(*
SPDX-FileCopyrightText: © 2026 Oleksandr Tiutyk <trofimich@gmail.com>
SPDX-License-Identifier: MIT
License: https://opensource.org/license/mit
*)

(*!
<summary>Concrete CatchActivity implementation for testing TryCatch exception capture and recovery.</summary>
*)

{attribute 'no_explicit_call' := 'do not call this function block directly'}
{attribute 'enable_dynamic_creation'}
FUNCTION_BLOCK RecoveryCatchTestActivity EXTENDS TOF_Workflow.CatchActivity
VAR_STAT
	{attribute 'hide'}
	_RecoveryCatchClassName : STRING := __POUNAME();
END_VAR
VAR
	_Recovered : BOOL;
END_VAR

//! <summary>Borrows the concrete class name for the lifetime of this instance.</summary>
{attribute 'monitoring' := 'call'}
PROPERTY ClassName : REFERENCE TO STRING
GET
ClassName REF= _RecoveryCatchClassName;
END_GET
END_PROPERTY

{attribute 'monitoring' := 'call'}
PROPERTY NamespaceName : REFERENCE TO STRING
GET
NamespaceName REF= CurrentNamespace.Name;
END_GET
END_PROPERTY

METHOD PROTECTED OnRunning : TOF_Workflow.ACTIVITY_RUNNING_STATE
VAR_INPUT
	startRunning : BOOL;
	startResuming : BOOL;
END_VAR
VAR_OUTPUT
	haltReason : WSTRING(255);
END_VAR
VAR
	variableFound : BOOL;
	errorHandledVar : TOF_Core.GENERIC_VALUE;
	trueValue : BOOL := TRUE;
END_VAR
_Recovered := TRUE;

variableFound := TryGetVariable(name := 'ErrorHandled', variable => errorHandledVar);

IF variableFound THEN
	errorHandledVar.ChangeValueByAnyType(value := trueValue, isObject := FALSE);
END_IF

OnRunning := TOF_Workflow.ACTIVITY_RUNNING_STATE.WORK_COMPLETED;
END_METHOD

METHOD PROTECTED OnStopping : TOF_Workflow.ACTIVITY_STOPPING_STATE
VAR_INPUT
	startCancelling : BOOL;
	startSuspending : BOOL;
END_VAR
VAR_OUTPUT
	haltReason : WSTRING(255);
END_VAR
OnStopping := TOF_Workflow.ACTIVITY_STOPPING_STATE.WORK_STOPPED;
END_METHOD

PROPERTY Recovered : BOOL
GET
Recovered := _Recovered;
END_GET
END_PROPERTY

{attribute 'monitoring' := 'call'}
PROPERTY SelfSize : ULINT
GET
SelfSize := XSIZEOF(THIS^);
END_GET
END_PROPERTY

END_FUNCTION_BLOCK

(* stored: Version 1.1.0.1
   POU RecoveryCatchTestActivity: Id {9ef9cde4-4a42-4ce8-bb7c-9a980b08bccc}, SpecialFunc None
   Property ClassName: Id {1173b19f-9d96-45f0-afe2-773bd386ab7a}
   Get Get: Id {c9c9a1df-27a4-45f5-8aba-4d02cde36f5b}
   Property NamespaceName: Id {134a2567-5247-42c8-9c2a-d9cd426bc35e}
   Get Get: Id {e8f6db09-7587-4387-8e55-6fe1f0b42130}
   Method OnRunning: Id {e2bc463e-e145-4216-9f96-737e127dba3c}
   Method OnStopping: Id {bf8c39bc-02d6-4406-a786-f5a04b4d568f}
   Property Recovered: Id {3d14b445-b3e3-4a47-a045-23af0b665631}
   Get Get: Id {6e2b5aea-0c16-4791-b124-246c5ae5d044}
   Property SelfSize: Id {1b6f75d9-93b2-4e0e-b411-2608e1e2498f}
   Get Get: Id {f1973ea9-caf7-4e48-855f-ffdb09f3e7a4} *)
